//---------------------------------------------------------------------------------------------------------------
//
//  HAUD 2026.01.16
//
//  - ExternControl
//
//    - placeholder programm for specific implementation of machine logic
//
//---------------------------------------------------------------------------------------------------------------
PROGRAM MAIN
VAR
	bInit 				          : BOOL;
  eInit                   : E_PROGRESS := E_PROGRESS.PROGRESS_DONE; // empty right now, so init is done
END_VAR

//---------------------------------------------------------------------------------------------------------------
// VISU POOL
//  - collect data to display
//  - set commands to structures
//---------------------------------------------------------------------------------------------------------------
VISU_POOL();
//---------------------------------------------------------------------------------------------------------------
//---------------------------------------------------------------------------------------------------------------

END_PROGRAM

(* stored: Version 1.1.0.1
   POU MAIN: Id {45b4bab1-5ef6-4038-a1c1-76ecc634eeae}, SpecialFunc None *)
